(* IEC 61131-3 sources: FibonacciChallenge/Network, 1 file *)

(* ---- ConfigObjects.st ---- *)
FUNCTION GLOBAL TAB TASK_CONF
_K_TASK, _K_REAL,
_K_END_VAR,

_K_TASK, _K_CYCLIC,
_K_END_VAR,

_K_TASK, _K_BACKGROUND,
_K_END_VAR,

_K_END_CONF
END_FUNCTION

FUNCTION GLOBAL TAB IPR_CONF
_K_IPR
	0$UINT,
_K_END_VAR,
_K_END_CONF
END_FUNCTION

FUNCTION GLOBAL TAB CONFIG_TABLES
00055$UINT,
0$UINT, 0, 4, "_CAN",
0$UINT, 1, 10, "_CANLIB",
0$UINT, 1, 20, "_FILESYS",
0$UINT, 1, 1, "_MULTITASK",
0$UINT, 0, 5, "_OSKERNEL",
0$UINT, 1, 34, "_SERLIB",
0$UINT, 0, 0, "_STDLIB",
0$UINT, 1, 1, "_TASKOBJECTCONTROL",
0$UINT, 1, 21, "ASCII_BIN",
0$UINT, 1, 24, "BUSINTERFACESDIAS",
0$UINT, 2, 0, "BUSINTERFACESDIASINTERNAL",
0$UINT, 1, 1, "CP112_IOS",
0$UINT, 0, 4, "CRITICALSECTION",
0$UINT, 2, 33, "DIASMASTER",
0$UINT, 1, 82, "DIASMASTERC",
0$UINT, 2, 24, "DIASMASTERMAIN",
0$UINT, 1, 0, "DIASMASTERPOSTSCAN",
0$UINT, 1, 14, "DM161",
0$UINT, 1, 11, "EEPROM",
0$UINT, 0, 0, "FIBCHALLENGE",
0$UINT, 1, 21, "HUB_BASE",
0$UINT, 2, 11, "HUB_BASE_ROOT",
0$UINT, 2, 35, "HWBASE",
0$UINT, 2, 55, "HWBASECDIAS",
0$UINT, 1, 0, "HWCLOGGING",
0$UINT, 5, 14, "HWCONTROL",
0$UINT, 1, 10, "HWCONTROLBASE",
0$UINT, 1, 0, "HWRTPOSTSCAN",
0$UINT, 1, 6, "I2CCDIAS",
0$UINT, 1, 22, "MERKEREX",
0$UINT, 0, 0, "MYFIRSTCLASS",
0$UINT, 1, 9, "RAMFILE",
0$UINT, 1, 24, "SAFETYBASEFSOE",
0$UINT, 3, 17, "SAFETYCDIAS_BASE",
0$UINT, 2, 18, "SAFETYMANAGER",
0$UINT, 1, 4, "SAFETYUDP",
0$UINT, 1, 37, "SCP111",
0$UINT, 1, 60, "SDIASBASE",
0$UINT, 1, 10, "SDIASHUBBASE",
0$UINT, 1, 94, "SDIASMANAGER",
0$UINT, 2, 3, "SDIASPLC",
0$UINT, 1, 9, "SDIASSAFETYBASE",
0$UINT, 1, 26, "SDIASSAFETYMANAGERFSOE",
0$UINT, 1, 11, "SDM081",
0$UINT, 0, 34, "SIGCLIB",
0$UINT, 1, 11, "STRING",
0$UINT, 1, 84, "STRINGINTERNAL",
0$UINT, 1, 21, "SYNCCALL",
0$UINT, 2, 17, "VARAN_BASE",
0$UINT, 3, 3, "VARANMANAGER",
0$UINT, 2, 4, "VARANMANAGER_1",
0$UINT, 1, 25, "VARANMANAGER_BASE",
0$UINT, 1, 3, "VIRTUALBASEINIT",
0$UINT, 2, 11, "WATCHDOGDIAS",
0$UINT, 1, 1, "XXXBASE_IOS",
ONE_CFG$UINT, 0, 0, "ONE_FibonacciChallegeNetwork",
TASK_CFG$UINT, 0, 0, "TASK_CONF",
IPR_CFG$UINT, 0, 0, "IPR_CONF",
PRJ_CFG$UINT, 0, 0, "FibChallenge",
END_FUNCTION

FUNCTION GLOBAL TAB CH_REDIRECT_EMB_TAB
0000$UINT,
00013$UINT,
"BUSINTERFACESDIAS;SERIALNO", "\SERIALNOSTR.DATA",
"DM161;SERIALNO", "\SERIALNOSTR.DATA",
"HWBASECDIAS;SERIALNO", "\SERIALNOSTR.DATA",
"SAFETYCDIAS_BASE;SERIALNO", "\SERIALNOSTR.DATA",
"SCP111;DESIGNERPRJNAME", "\SDIASSAFETYMANAGERFSOE1\PROJECTNAMESTR.DATA",
"SCP111;DESIGNERPRJREV", "\SDIASSAFETYMANAGERFSOE1\PROJECTREVISIONSTR.DATA",
"SCP111;SERIALNO", "\SERIALNOSTR.DATA",
"SDIASBASE;SERIALNO", "\SERIALNOSTR.DATA",
"SDIASSAFETYBASE;SERIALNO", "\SERIALNOSTR.DATA",
"SDIASSAFETYMANAGERFSOE;DESIGNERPRJNAME", "\PROJECTNAMESTR.DATA",
"SDIASSAFETYMANAGERFSOE;DESIGNERPRJREV", "\PROJECTREVISIONSTR.DATA",
"SDM081;SERIALNO", "\SERIALNOSTR.DATA",
"VARAN_BASE;SERIALNO", "\SERIALNOSTR.DATA",
END_FUNCTION
